Fanuc KAREL source: KB00128.KL

PROGRAM KB00128
%NOLOCKGROUP
%ENVIRONMENT VECTR
VAR
  P1: POSITION
  RESULT: VECTOR
BEGIN
  RESULT = ORIENT(P1)
END KB00128
